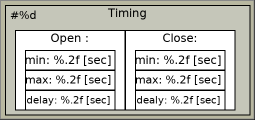
VISUALIZATION vis_Piston_Times  // 255x120
VAR_IN_OUT
	stPis: ST_Piston;
END_VAR
    Rectangle (0,0 255x120)
    Rectangle (5,5 245x110), "Timing"
    Rectangle (15,30 110x80), "Open :"
    Rectangle (125,30 110x80), "Close:"
    Rectangle (135,50 90x20), "min: %.2f [sec]", text variable: stPis.t_minClose
        OnMouseDown: write the text variable via Edit, min 0
    Rectangle (135,70 90x20), "max: %.2f [sec]", text variable: stPis.t_maxClose
        OnMouseDown: write the text variable via Edit, min 0
    Rectangle (25,70 90x20), "max: %.2f [sec]", text variable: stPis.t_maxOpen
        OnMouseDown: write the text variable via Edit, min 0
    Rectangle (25,50 90x20), "min: %.2f [sec]", text variable: stPis.t_minOpen
        OnMouseDown: write the text variable via Edit, min 0
    Rectangle (25,90 90x20), "delay: %.2f [sec]", text variable: stPis.t_DelayOpen
        OnMouseDown: write the text variable via Edit, min 0
    Rectangle (135,90 90x20), "dealy: %.2f [sec]", text variable: stPis.t_DelayClose
        OnMouseDown: write the text variable via Edit, min 0
    Textfield (4,5 39x21), "#%d", text variable: stPis.iPisNum
END_VISUALIZATION

(* stored: Version 1.1.0.1, ProductVersion 3.1.4024.12
   Visu vis_Piston_Times: Id {04fb3c0a-e576-4324-b930-54f0392269b4} *)
